(*
SPDX-FileCopyrightText: © 2026 Oleksandr Tiutyk <trofimich@gmail.com>
SPDX-License-Identifier: MIT
License: https://opensource.org/license/mit
*)

(*!
<summary>Provides a test exception whose GetMessage deliberately throws another exception.</summary>
<description>
Static Throw clones this concrete type. The clone is task-managed; GetMessage deliberately throws a separate
StandardException. The per-instance call count records formatter invocations and is independent of diagnostic
payload. This fixture never performs I/O or throws from lifecycle initialization.
</description>
*)

{attribute 'enable_dynamic_creation'}
FUNCTION_BLOCK ThrowingGetMessageException EXTENDS TOF_Core.StandardException
VAR
	_FixtureClassName : STRING := __POUNAME();
	_MessageReadCount : UDINT;
END_VAR

{attribute 'monitoring' := 'call'}
PROPERTY ClassName : REFERENCE TO STRING
GET
ClassName REF= _FixtureClassName;
END_GET
END_PROPERTY

(*!
<summary>Creates a task-managed clone retaining the failing formatter.</summary>
<description>
Registers the new object before copying inherited diagnostics. Its formatter invocation count starts at zero.
The caller borrows the result until task cleanup. Allocation failure follows the framework terminal policy.
</description>
*)
METHOD Clone : TOF_Core.IObject
VAR
	copy : POINTER TO ThrowingGetMessageException;
END_VAR
copy := __NEW(ThrowingGetMessageException);

IF copy = 0 THEN
	TOF_Core.DynamicMemoryManager.RaiseAllocationFailure();
END_IF

TOF_Core.DynamicMemoryManager.RegisterAutoDisposedObject(autoDisposedObject := copy^);
copy^.CopyGeneralFields(sourceException := THIS^);
Clone := copy^;
END_METHOD

(*!
<summary>Deliberately fails while formatting the original child exception.</summary>
<description>
Counts the call before throwing so tests can distinguish formatter failure from early refusal.
Neither formatting option is used.
</description>
<param name="showSource">Unused formatting option retained for the inherited signature.</param>
<param name="timestampDisplayMode">Unused formatting option retained for the inherited signature.</param>
*)
METHOD GetMessage : TOF_Core.ERROR_MESSAGE
VAR_INPUT
	showSource : BOOL := FALSE;
	timestampDisplayMode : TOF_Core.TIMESTAMP_DISPLAY_MODE := TOF_Core.TIMESTAMP_DISPLAY_MODE.HIDDEN;
END_VAR
VAR
	failure : TOF_Core.StandardException;
END_VAR
_MessageReadCount := _MessageReadCount + 1;

failure.Throw(
	sourceNamespaceName := NamespaceName,
	sourceClassName := ClassName,
	sourcePOUName := __POUNAME(),
	sourcePosition := __POSITION(),
	message := "Injected message formatting failure"
);
END_METHOD

(*!
<summary>Borrows the test library namespace.</summary>
*)

{attribute 'monitoring' := 'call'}
PROPERTY NamespaceName : REFERENCE TO STRING
GET
NamespaceName REF= CurrentNamespace.Name;
END_GET
END_PROPERTY

(*!
<summary>Reports the concrete fixture size.</summary>
*)

{attribute 'monitoring' := 'call'}
PROPERTY SelfSize : ULINT
GET
SelfSize := XSIZEOF(THIS^);
END_GET
END_PROPERTY

//! <summary>Counts this instance's formatter calls, including ones that raised the injected exception.</summary>
PROPERTY MessageReadCount : UDINT
GET
MessageReadCount := _MessageReadCount;
END_GET
END_PROPERTY

END_FUNCTION_BLOCK

(* stored: Version 1.1.0.1, ProductVersion 3.1.4026.21
   POU ThrowingGetMessageException: Id {b209960a-a1ef-448b-a416-34bdbbe0f5b1}, SpecialFunc None
   Property ClassName: Id {335aa07b-233f-4826-9c68-97ff972abb42}
   Get Get: Id {07fa6a19-5bcb-464d-a105-d1aa193d86bb}
   Method Clone: Id {ded3acc1-405f-42bb-8bea-1304bbdc3356}
   Method GetMessage: Id {5bf4a784-1969-4915-94b1-50b5d93ff030}
   Property NamespaceName: Id {534173d0-7c8b-442e-92ad-0a298013a260}
   Get Get: Id {53c744f6-bf11-4262-89c6-e2b4f467b8b5}
   Property SelfSize: Id {e460b78a-3e7a-45e0-a978-d398889a0791}
   Get Get: Id {af579f54-2ae9-48d2-8882-fa728cfb3c77}
   Property MessageReadCount: Id {8ac09787-ffcb-4777-b5e6-53940df01a83}
   Get Get: Id {d21dc32e-1c6a-4778-ac5e-c30e3e68e849} *)
